(* IEC 61131-3 sources: sis-interlock-demo/src/POUs/Sis/F_SisAiToEu, 1 file *)

(* ---- F_SisAiToEu.decl.st ---- *)
// Назначение: ток 4–20 мА в инженерные единицы по шкале датчика, без ограничения: выход за
//             шкалу сохраняется, недостоверность решает F_SisNe43Valid.
// Автор:      kr0nsch
// Версия:     0.1.0
// Документ:   docs/DESIGN.md, раздел «8.3 Аналоговые входы 4–20 мА (NE 43)»
// ВНИМАНИЕ:   код демонстрационный и не предназначен для систем безопасности. Реальная ПАЗ
//             требует определения SIL, сертифицированных аппаратных и программных средств
//             и валидации по ГОСТ Р МЭК 61511.
FUNCTION F_SisAiToEu : REAL
VAR_INPUT
    rIn_mA : REAL;   // ток канала, мА
    rLo_eu : REAL;   // значение при 4 мА, инж. ед.
    rHi_eu : REAL;   // значение при 20 мА, инж. ед.
END_VAR
